TYPE ST_Pump :
STRUCT
	//request
	modeAuto	:	BOOL	;//System in automatic
	bRun_Auto	:	BOOL	;
	bRun_Man	:	BOOL	;
	bRun		: 	BOOL;
	DriveReady	: 	BOOL;

	nRPM_Auto	:	REAL		;//Pump RPM 
	nRPM_Man	:	REAL		;//Pump RPM 
	nRPM		:	REAL		;//Pump RPM 
	//feedback
	nRPM_fdbk	:	INT	;
END_STRUCT
END_TYPE

(* stored: Version 1.1.0.1, ProductVersion 3.1.4024.13
   DUT ST_Pump: Id {2d6d8fa6-e575-4761-89fb-cc0bf15c71a5} *)
